ABB RAPID module: user.sys

MODULE user (SYSMODULE)

 ! Predefined user data
 !*********************

 ! Declaration of numeric registers reg1...reg5
 VAR num reg1 := 0;
 VAR num reg2 := 0;
 VAR num reg3 := 0;
 VAR num reg4 := 0;
 VAR num reg5 := 0;

 ! Declaration of stopwatch clock1
 VAR clock clock1;

 ! Template for declaration of workobject wobj1
 !TASK PERS wobjdata wobj1 := [FALSE, TRUE, "", [[0, 0, 0],[1, 0, 0, 0]],[[0, 0, 0],[1, 0, 0, 0]]];

ENDMODULE
